(* IEC 61131-3 sources: codesys-to-astra/corpus/boiler-plc210/src/GVLs, 5 files *)

(* ---- GVL_Clock.gvl.st ---- *)
// Назначение: время ПЛК из каналов узла OwenRTC и данные узла Watchdog.
// Автор:      kr0nsch
// Версия:     0.1.0
// Документ:   corpus/boiler-plc210/README.md
VAR_GLOBAL
    dtNow : DT;             // Date And Time
    sDateText : STRING(80); // Format date
    sTimeText : STRING(80); // Format time
    usiHour : USINT;        // Hour
    usiWeek : USINT;        // Week of year
    udiLastExc : UDINT;     // Watchdog: код последнего исключения
END_VAR

(* ---- GVL_Hmi.gvl.st ---- *)
// Назначение: строки и коды для панели оператора.
// Автор:      kr0nsch
// Версия:     0.1.0
// Документ:   corpus/boiler-plc210/README.md
VAR_GLOBAL
    sStatus : STRING(255);  // строка состояния
    sCode : STRING(8);      // код состояния (hex)
    eState : E_BoilerState; // состояние котла К1
END_VAR

(* ---- GVL_Hw.gvl.st ---- *)
// Назначение: встроенный ввод-вывод ПЛК210 по AT-адресам (так делать ОВЕН не рекомендует — Targets v3.4, разд. 1;
//             вход нарочно с AT, чтобы показать C2A-IO001).
// Автор:      kr0nsch
// Версия:     0.1.0
// Документ:   corpus/boiler-plc210/README.md
VAR_GLOBAL
    xBurner1Fault AT %IX0.0 : BOOL;     // авария горелки К1
    xBurner2Fault AT %IX0.1 : BOOL;     // авария горелки К2
    xPumpRun AT %QX0.0 : BOOL;          // пуск сетевого насоса Н1
    xAlarmHorn AT %QX0.1 : BOOL;        // сирена
    wHmiStatus AT %MW10 : WORD;         // слово состояния для панели
END_VAR

(* ---- GVL_Mx.gvl.st ---- *)
// Назначение: значения модулей Mx210 (привязки к каналам шаблонов МВ210-101 и МУ210-402 в дереве устройств).
// Автор:      kr0nsch
// Версия:     0.1.0
// Документ:   corpus/boiler-plc210/README.md
VAR_GLOBAL
    rTSupply_C : REAL;      // температура подачи, °C (МВ210-101, вход 1)
    rTReturn_C : REAL;      // температура обратки, °C (вход 2)
    rTOutdoor_C : REAL;     // температура наружного воздуха, °C (вход 3)
    iTSupplyRaw : INT;      // подача, целое (вход 1, integer)
    wDoMask : WORD;         // выходы МУ210-402 (битовая маска)
    wMeterStatus : WORD;    // счётчик энергии на Modbus 3S (канал FC 23)
END_VAR

(* ---- GVL_Persist.gvl.st ---- *)
// Назначение: сохраняемые уставки и наработка.
// Автор:      kr0nsch
// Версия:     0.1.0
// Документ:   corpus/boiler-plc210/README.md
VAR_GLOBAL RETAIN
    rSpBase_C : REAL := 70.0;   // базовая уставка подачи, °C
    udiRunTime_s : UDINT;       // наработка насоса, с
END_VAR
